// TIA Portal project "Ligne_auto" (V16)

(* hardware
DEVICE "Station S7300/ET200M_1"  S7-300 station
   slot 0: "Châssis_0"  Rail  6ES7 390-1***0-0AA0
   slot 2: "PLC_1"  CPU 314C-2 PN/DP  6ES7 314-6EH04-0AB0  V3.3
      slot 2: "Interface PROFINET_1"  PN-IO
         slot 1: "Port_1"  Port
         slot 2: "Port_2"  Port
      slot 5: "DI 24/DO 16_1"  DI24/DO16
      slot 6: "AI 5/AO 2_1"  AI5/AO2
      slot 7: "Comptage_1"  Counter
      slot 8: "Positionnement_1"  Positioning
*)

// ===== PLC "PLC_1"  CPU 314C-2 PN/DP =====

VAR_GLOBAL   // PLC tag table "Table de variables standard"
   "BP_MARCHE" AT %I0.0 : Bool;
   "BP_ARRET" AT %I0.1 : Bool;
   "ARRET_URGENCE_OK" AT %I0.2 : Bool;
   "PRESENCE_ENTREE" AT %I0.3 : Bool;
   "PRESENCE_CONTROLE" AT %I0.4 : Bool;
   "CAPTEUR_METAL" AT %I0.5 : Bool;
   "CAPTEUR_HAUTEUR" AT %I0.6 : Bool;
   "PIECE_BAC1" AT %I0.7 : Bool;
   "PIECE_BAC2" AT %I1.0 : Bool;
   "PIECE_BAC3" AT %I1.1 : Bool;
   "AIGUILLAGE_REPOS" AT %I1.2 : Bool;
   "DEFAUT_MOTEUR" AT %I1.3 : Bool;
   "BP_REARMEMENT" AT %I1.4 : Bool;
   "MOTEUR_CONVOYEUR" AT %Q0.0 : Bool;
   "TRI_BAC1" AT %Q0.1 : Bool;
   "TRI_BAC2" AT %Q0.2 : Bool;
   "TRI_BAC3" AT %Q0.3 : Bool;
   "VOYANT_MARCHE" AT %Q0.4 : Bool;
   "VOYANT_DEFAUT" AT %Q0.5 : Bool;
   "BUZZER" AT %Q0.6 : Bool;
   "VOYANT_ARRET" AT %Q0.7 : Bool;
END_VAR

FUNCTION_BLOCK "GFN"   // FB1, GRAPH
{ S7_Optimized_Access := 'FALSE' }
VERSION : 0.1
   VAR_INPUT
      OFF_SQ : Bool := false;   // Désactiver le graphe
      INIT_SQ : Bool := false;   // Mettre le graphe à l'état initial
      ACK_EF : Bool := false;   // Acquitter toutes les erreurs et perturbations
      S_PREV : Bool := false;   // Afficher l'étape précédente dans le paramètre S_NO
      S_NEXT : Bool := false;   // Afficher l'étape suivante dans le paramètre S_NO
      SW_AUTO : Bool := false;   // Mode automatique
      SW_TAP : Bool := false;   // Mode semi-automatique/Activation de l'étape suivante avec transition
      SW_TOP : Bool := false;   // Mode semi-automatique/Ignorer la transition
      SW_MAN : Bool := false;   // Mode manuel
      S_SEL : Int := 0;   // Sélectionner l'étape à afficher dans S_NO
      S_ON : Bool := false;   // Activer l'étape figurant dans le paramètre S_NO
      S_OFF : Bool := false;   // Désactiver l'étape figurant dans le paramètre S_NO
      T_PUSH : Bool := false;   // Validation de commutation pour transition en mode semi-automatique
   END_VAR
   VAR_OUTPUT
      S_NO : Int := 0;   // Numéro d'étape
      S_MORE : Bool := false;   // Il existe d'autres étapes qui peuvent être affichées dans S_NO.
      S_ACTIVE : Bool := false;   // L'étape affichée dans le paramètre S_NO est activée
      ERR_FLT : Bool := false;   // Erreur groupée Interlock or Supervision
      AUTO_ON : Bool := false;   // Mode automatique activé
      TAP_ON : Bool := false;   // Mode semi-automatique/Etape avec transition activé
      TOP_ON : Bool := false;   // Mode semi-automatique/Ignorer la transition activé
      MAN_ON : Bool := false;   // Mode manuel activé
   END_VAR
   VAR
      S_DISPLAY : Int;   // Affichage interne du paramètre de sortie S_NO
      S_SEL_OLD : Int;   // Valeur précédente dans S_SEL
      S_DISPIDX : Byte;   // Indice de l'étape affichée dans S_NO
      T_DISPIDX : Byte;   // Indice de la transition affichée dans T_NO
      MOP : Struct   // Mode de fonctionnement
         AUTO : Bool := true;   // Etat : Mode automatique
         MAN : Bool := false;   // Etat : Mode manuel
         TAP : Bool := false;   // Etat : Mode semi-automatique/Activation de l'étape suivante avec transition
         TOP : Bool := false;   // Etat : Mode semi-automatique/Ignorer la transition
         ACK_S : Bool := false;   // Requête : Acquitter l'étape figurant dans le paramètre S_NO
         REG_S : Bool := false;   // Requête : Enregistrer l'étape figurant dans le paramètre S_NO
         T_PREV : Bool := false;   // Requête : Afficher la transition valide précédente dans le paramètre T_NO
         T_NEXT : Bool := false;   // Requête : Afficher la transition valide suivante dans le paramètre T_NO
         LOCK : Bool := true;   // Etat : Traitement des Interlocks activé
         SUP : Bool := true;   // Etat : Traitement de Supervision activé
         ACKREQ : Bool := true;   // Etat : Acquittement requis
         SSKIP : Bool := false;   // Etat : "Ignorer les étapes" activé
         OFF : Bool := false;   // Requête : Désactiver toutes les étapes
         INIT : Bool := true;   // Requête : Mettre le graphe à l'état initial
         HALT : Bool := false;   // Etat : Le graphe est arrêté
         TMS_HALT : Bool := false;   // Etat : Toutes les temporisations internes sont arrêtées
         OPS_ZERO : Bool := false;   // Etat : Tous les opérandes traités avec N, L, D mis à 0
         SACT_DISP : Bool := true;   // Etat : N'afficher que les étapes actives
         SEF_DISP : Bool := false;   // Etat : Afficher uniquement les étapes avec erreurs et perturbations
         SALL_DISP : Bool := false;   // Etat : Afficher toutes les étapes
         S_PREV : Bool := false;   // Requête : Afficher l'étape précédente dans le paramètre S_NO
         S_NEXT : Bool := false;   // Requête : Afficher l'étape suivante dans le paramètre S_NO
         S_SELOK : Bool := false;   // Requête : Afficher dans le paramètre S_NO le numéro d'étape figurant dans S_SEL
         S_ON : Bool := false;   // Requête : Activer l'étape figurant dans le paramètre S_NO
         S_OFF : Bool := false;   // Requête : Désactiver l'étape figurant dans le paramètre S_NO
         T_PUSH : Bool := false;   // Requête : Validation de commutation pour transition
         REG : Bool := false;   // Requête : Enregistrer toutes les erreurs Interlock et Supervision
         ACK : Bool := false;   // Requête : Acquitter toutes les erreurs Interlock et Supervision
         IL_PERM : Bool := false;   // Etat : Traitement permanent de tous les Interlocks
         T_PERM : Bool := false;   // Etat : Traitement permanent de toutes les transitions
         ILP_MAN : Bool := false;   // Etat : Traitement permanent de tous les Interlocks en mode manuel
      END_STRUCT;
      TICKS : Struct   // Périodes d'horloge
         DELTA : Time := T#0ms;   // Différence de temps entre deux cycles
         OLD : Time := T#0ms;   // Valeur du compteur de périodes 10 ms au dernier cycle
         NEW : Time := T#0ms;   // Valeur du compteur de périodes 10 ms dans ce cycle
      END_STRUCT;
      SQ_FLAGS : Struct   // Mémentos de graphe
         ERR_FLT : Bool := false;   // Erreur groupée Interlock et Supervision
         ERROR : Bool := false;   // Erreur groupée Interlock
         FAULT : Bool := false;   // Erreur groupée Supervision
         RT_FAIL : Bool := false;   // Erreur à l'exécution
         NO_SNO : Bool := false;   // Numéro d'étape requis introuvable
         NF_OFL : Bool := false;   // Débordement : Trop de requêtes ON ou OFF
         SA_OFL : Bool := false;   // Débordement : Trop d'étapes activées
         TV_OFL : Bool := false;   // Débordement : Trop de transitions valides
         MSG_OFL : Bool := false;   // Débordement : Pas assez de ressources système pour ALARM_S
         NO_SWI : Bool := false;   // Pas de commutation dans ce cycle
         CYC_OP : Bool := false;   // Exécution cyclique du graphe après l'initialisation
         AS_MSG : Bool := true;   // Messages à l'exécution activés ou désactivés par instruction
         AS_SEND : Bool := false;   // Envoyer les messages de WR_USMSG ou les entrer uniquement dans le tampon de diagnostic
         SQ_BUSY : Bool := false;   // Mémento de front interne pour le traitement séquentiel
         SA_BUSY : Bool := false;   // Mémento de front interne pour le traitement séquentiel
         AS_SIG : Bool := false;   // Mémentos de front pour messages de Alarm_S et Alarm_SQ
      END_STRUCT;
   END_VAR
BEGIN
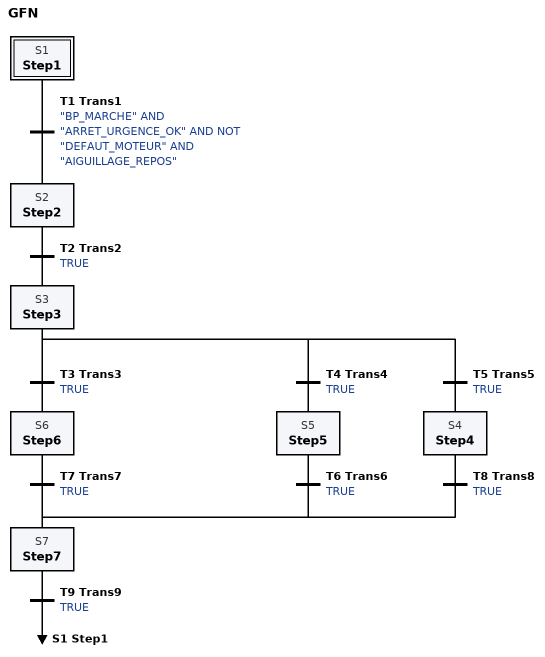
   // sequencer 1
   INITIAL_STEP Step1:   // S1
   END_STEP
   TRANSITION Trans1 FROM Step1 TO Step2   // T1
      := "BP_MARCHE" AND "ARRET_URGENCE_OK" AND NOT "DEFAUT_MOTEUR" AND "AIGUILLAGE_REPOS";
   END_TRANSITION
   STEP Step2:   // S2
   END_STEP
   TRANSITION Trans2 FROM Step2 TO Step3   // T2
      := TRUE;
   END_TRANSITION
   STEP Step3:   // S3
   END_STEP
   TRANSITION Trans3 FROM Step3 TO Step6   // T3
      := TRUE;
   END_TRANSITION
   TRANSITION Trans4 FROM Step3 TO Step5   // T4
      := TRUE;
   END_TRANSITION
   TRANSITION Trans5 FROM Step3 TO Step4   // T5
      := TRUE;
   END_TRANSITION
   STEP Step4:   // S4
   END_STEP
   TRANSITION Trans8 FROM Step4 TO Step7   // T8
      := TRUE;
   END_TRANSITION
   STEP Step5:   // S5
   END_STEP
   TRANSITION Trans6 FROM Step5 TO Step7   // T6
      := TRUE;
   END_TRANSITION
   STEP Step6:   // S6
   END_STEP
   TRANSITION Trans7 FROM Step6 TO Step7   // T7
      := TRUE;
   END_TRANSITION
   STEP Step7:   // S7
   END_STEP
   TRANSITION Trans9 FROM Step7 TO Step1   // T9, jump
      := TRUE;
   END_TRANSITION
END_FUNCTION_BLOCK

ORGANIZATION_BLOCK "Main"   // OB1, LAD
TITLE = "Main Program Sweep (Cycle)"
{ S7_Optimized_Access := 'FALSE' }
VERSION : 0.1
   VAR_TEMP
      OB1_EV_CLASS : Byte;   // Bits 0-3 = 1 (Coming event), Bits 4-7 = 1 (Event class 1)
      OB1_SCAN_1 : Byte;   // 1 (Cold restart scan 1 of OB 1), 3 (Scan 2-n of OB 1)
      OB1_PRIORITY : Byte;   // Priority of OB Execution
      OB1_OB_NUMBR : Byte;   // 1 (Organization block 1, OB1)
      OB1_RESERVED_1 : Byte;   // Reserved for system
      OB1_RESERVED_2 : Byte;   // Reserved for system
      OB1_PREV_CYCLE : Int;   // Cycle time of previous OB1 scan (milliseconds)
      OB1_MIN_CYCLE : Int;   // Minimum cycle time of OB1 (milliseconds)
      OB1_MAX_CYCLE : Int;   // Maximum cycle time of OB1 (milliseconds)
      OB1_DATE_TIME : Date_And_Time;   // Date and time OB1 started
   END_VAR
BEGIN
END_ORGANIZATION_BLOCK